FUNCTION_BLOCK NctGripper EXTENDS CyclicComponent IMPLEMENTS I_NctGripper
VAR
	_DwellTimer			: TON; //Q = the gripper has held the last output change for _ActionTime
	_ActionTime			: TIME	:= T#10MS; //Minimum time the gripper holds each output state; it takes one command per 10 ms
	_OpenPosition		: LREAL := 0.05;
	_ClosePosition		: LREAL := 9.3;
	_Simulated			: BOOL;
	_SimActionTime		: TIME;
	_SimTimer			: TON;
	_NctBaseUnit		: I_XtsNctBaseUnit;
	_GripperOpen		: NctDigitalOutput('Gripper Open', 1);
	_GripperClose		: NctDigitalOutput('Gripper Close', 3);
	_GripperPos			: NctAnalogInput('Gripper Position', 1);
	_OutputChangeCount	: UDINT; //ProcessDataUpdateCount when an output last changed
	_PowerUpTime		: TIME	:= T#30MS; //Exchanges must have run this long before a pulse starts; the gripper ignores an input that is already on when it powers up
	_PowerUpTimer		: TON; //Q = on an NCT module and powered up for _PowerUpTime
	_NoExchangeTimer	: TON; //Q = no NCT exchange for 30 ms, the mover is off the module
	_LastUpdateCount	: UDINT;
END_VAR

METHOD Close : BOOL
IF _GripperClose.On THEN
	Close := TRUE; //Pulse already running
	RETURN;
END_IF

//Only start on a powered-up module, after any Open pulse has ended and the all-off state has been held
IF _GripperOpen.On OR NOT _PowerUpTimer.Q OR NOT _DwellTimer.Q THEN
	RETURN;
END_IF

SetOutputs(OpenOn := FALSE, CloseOn := TRUE);
Close := TRUE;
END_METHOD

PROPERTY CloseOutput : I_DigitalOutput
GET
CloseOutput := _GripperClose;
END_GET
END_PROPERTY

METHOD CyclicLogic
//The gripper only has power on an NCT module, and ignores an input that is already on when it powers up
_NoExchangeTimer(IN := _NctBaseUnit.ProcessDataUpdateCount = _LastUpdateCount, PT := T#30MS);
_LastUpdateCount := _NctBaseUnit.ProcessDataUpdateCount;
_PowerUpTimer(IN := _Simulated OR NOT _NoExchangeTimer.Q, PT := _PowerUpTime);
IF NOT _PowerUpTimer.IN THEN
	SetOutputs(OpenOn := FALSE, CloseOn := FALSE); //Drop the command rather than deliver it at power-up
END_IF

//The gripper only sees the output image once per NCT exchange, so the hold starts when the mover acknowledges the change
_DwellTimer(IN := _Simulated OR ExchangesSinceChange() >= 2, PT := _ActionTime);
IF (_GripperOpen.On OR _GripperClose.On) AND _DwellTimer.Q THEN
	SetOutputs(OpenOn := FALSE, CloseOn := FALSE);
END_IF

_SimTimer(IN := _Simulated AND (_GripperOpen.On OR _GripperClose.On OR _SimTimer.IN), PT := _SimActionTime);
//Need to fix since changing to NCTAnalogInput
// IF _SimTimer.Q THEN
// 	IF _GripperPosition.Value <= _OpenPosition THEN
// 		_GripperPosition.ForceValue := LREAL_TO_INT(_ClosePosition);
// 	ELSE
// 		_GripperPosition.ForceValue := LREAL_TO_INT(_OpenPosition);
// 	END_IF
// END_IF
END_METHOD

//Completed NCT exchanges since an output last changed. 2 = the mover has acknowledged the frame carrying the change
METHOD PRIVATE ExchangesSinceChange : UDINT
ExchangesSinceChange := _NctBaseUnit.ProcessDataUpdateCount - _OutputChangeCount;
END_METHOD

(*FB_Init is always available implicitly and it is used primarily for initialization.
The return value is not evaluated. For a specific influence, you can also declare the
methods explicitly and provide additional code there with the standard initialization
code. You can evaluate the return value.*)
METHOD FB_Init : BOOL
VAR_INPUT
	(* TRUE: the retain variables are initialized (reset warm / reset cold)*)
	bInitRetains : BOOL;

	(* TRUE: the instance will be copied to the copy code afterward (online change)   *)
	bInCopyCode : BOOL;
	Name		: ApplicationBase.T_MaxString;
END_VAR
END_METHOD

{attribute 'monitoring' := 'call'}
PROPERTY GripperPosition : LREAL
GET
GripperPosition := _GripperPos.Value;
END_GET
END_PROPERTY

{attribute 'monitoring' := 'call'}
PROPERTY IsClosed : BOOL
GET
IsClosed := _GripperPos.Value > _ClosePosition;
END_GET
END_PROPERTY

{attribute 'monitoring' := 'call'}
PROPERTY IsOpen : BOOL
GET
IsOpen := _GripperPos.Value < _OpenPosition;
END_GET
END_PROPERTY

PROPERTY NctBaseUnit : I_XtsNctBaseUnit
GET
NctBaseUnit := _NctBaseUnit;
END_GET
SET
_NctBaseUnit			  := NctBaseUnit;
_GripperOpen.NctBaseUnit  := _NctBaseUnit;
_GripperClose.NctBaseUnit := _NctBaseUnit;
_GripperPos.NctBaseUnit	  := _NctBaseUnit;
END_SET
END_PROPERTY

METHOD Open : BOOL
IF _GripperOpen.On THEN
	Open := TRUE; //Pulse already running
	RETURN;
END_IF

//Only start on a powered-up module, after any Close pulse has ended and the all-off state has been held
IF _GripperClose.On OR NOT _PowerUpTimer.Q OR NOT _DwellTimer.Q THEN
	RETURN;
END_IF

SetOutputs(OpenOn := TRUE, CloseOn := FALSE);
Open := TRUE;
END_METHOD

PROPERTY OpenOutput : I_DigitalOutput
GET
OpenOutput := _GripperOpen;
END_GET
END_PROPERTY

PROPERTY PositionInput : I_AnalogInput
GET
PositionInput := _GripperPos;
END_GET
END_PROPERTY

METHOD PRIVATE SetOutputs
VAR_INPUT
	OpenOn	: BOOL;
	CloseOn : BOOL;
END_VAR
IF OpenOn AND CloseOn THEN
	RETURN; //The gripper rejects a command with both inputs on
END_IF

IF OpenOn <> _GripperOpen.On OR CloseOn <> _GripperClose.On THEN
	_GripperOpen.On	   := OpenOn;
	_GripperClose.On   := CloseOn;
	_OutputChangeCount := _NctBaseUnit.ProcessDataUpdateCount;
	_DwellTimer(IN := FALSE); //Restart the hold, and block another change in this same scan
END_IF
END_METHOD

{attribute 'monitoring' := 'call'}
PROPERTY Simulated : BOOL
GET
Simulated := _Simulated;
END_GET
SET
_Simulated := Simulated;

IF _Simulated THEN
	_GripperPos.Force := E_ForceState.ForceOn;
ELSE
	_GripperPos.Force := E_ForceState.Unforced;
END_IF
END_SET
END_PROPERTY

END_FUNCTION_BLOCK

(* stored: Version 1.1.0.1, ProductVersion 3.1.4026.21
   POU NctGripper: Id {63a0fe2a-ecd0-41f9-85f3-c919fae0008b}, SpecialFunc None
   Folder Constructor: Id {1a7e2c21-0bdc-49e3-a4ca-be3a4e537dc1}
   Folder Methods: Id {b69dec76-3681-4a6f-96b5-d6ec7a728651}
   Folder Properties: Id {00981d39-e99f-48e6-8097-b01b3e0a64e2}
   Method Close: Id {c9b47b51-4a28-43c6-8b4e-7c5fe527dc1d}
   Property CloseOutput: Id {c67c72d2-ea8e-47bd-9856-65b5f77423a3}
   Get Get: Id {f2b19d58-3e96-45f2-820b-3669a336d7cb}
   Method CyclicLogic: Id {f4e14436-77b9-4314-a73e-9057e2d853b8}
   Method ExchangesSinceChange: Id {79e030ca-6423-454a-891f-223b8989776d}
   Method FB_Init: Id {9023a8e8-1136-4d5b-9556-911beb55dac5}
   Property GripperPosition: Id {22a95f05-1a67-484c-a307-e5aec44ea7b4}
   Get Get: Id {1aa57a25-4ae2-4599-bf1e-1439ebb07bbe}
   Property IsClosed: Id {e485316b-bff0-468d-a813-b7c68e6d15d7}
   Get Get: Id {5a80ca39-986c-4e37-94aa-477d9e7de6d1}
   Property IsOpen: Id {254a9b7d-c468-4e24-a96c-ce0045de4085}
   Get Get: Id {981c13e7-62d3-4cd8-8f3e-139c8039e469}
   Property NctBaseUnit: Id {95a5f417-54ee-40ad-8435-a5d9e3783774}
   Get Get: Id {b22a6a00-5705-4231-a768-1e67277815c7}
   Set Set: Id {f74cde18-97c4-4f0c-ae71-adb1286c0b7c}
   Method Open: Id {692bc559-4382-47e8-97d6-0cfb3233bbbc}
   Property OpenOutput: Id {981fa11a-5cb1-4d21-94fc-2bf841550c06}
   Get Get: Id {4f16c2a1-b745-42ed-9abe-cee29af85d15}
   Property PositionInput: Id {75a14e3f-9819-49a5-abeb-00e2492bfa0e}
   Get Get: Id {d5ddf1c4-8cb9-4ee7-83d2-f0fef88415c8}
   Method SetOutputs: Id {236eb0fc-58e0-450c-ac4b-9e611d03cf35}
   Property Simulated: Id {e55fff7a-bccb-4a3e-a2ab-d1de12b96367}
   Get Get: Id {21da5f25-3753-4f87-8737-5b6e4d859c48}
   Set Set: Id {a33da3a8-aaab-474e-8261-7d02abe81fce} *)
